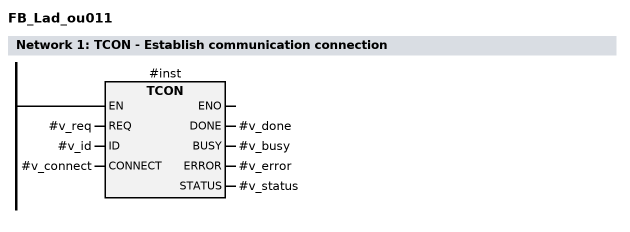
   #inst(REQ := #v_req,   // TCON
         ID := #v_id,
         CONNECT := #v_connect,
         DONE => #v_done,
         BUSY => #v_busy,
         ERROR => #v_error,
         STATUS => #v_status);
END_REGION
END_FUNCTION_BLOCK

FUNCTION_BLOCK "FB_Lad_ou012"   // FB78, LAD
{ S7_Optimized_Access := 'TRUE' }
   VAR_INPUT
      v_req : Bool;
      v_id : Word;
   END_VAR
   VAR_OUTPUT
      v_done : Bool;
      v_busy : Bool;
      v_error : Bool;
      v_status : Word;
   END_VAR
   VAR
      inst : TDISCON;
   END_VAR
BEGIN

REGION Network 1: TDISCON - Terminate communication connection
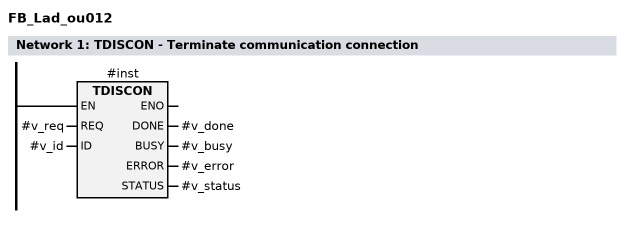
   #inst(REQ := #v_req, ID := #v_id, DONE => #v_done, BUSY => #v_busy, ERROR => #v_error, STATUS => #v_status);   // TDISCON
END_REGION
END_FUNCTION_BLOCK

FUNCTION_BLOCK "FB_Lad_ou013"   // FB79, LAD
{ S7_Optimized_Access := 'TRUE' }
   VAR_INPUT
      v_req : Bool;
      v_id : Conn_Ouc;
      v_len : UInt;
   END_VAR
   VAR_OUTPUT
      v_done : Bool;
      v_busy : Bool;
      v_error : Bool;
      v_status : Word;
   END_VAR
   VAR_IN_OUT
      v_data : Array[0..99] of Byte;
   END_VAR
   VAR
      inst : TSEND;
   END_VAR
BEGIN

REGION Network 1: TSEND - Send data via communication connection
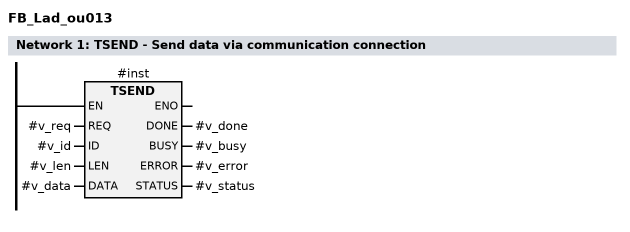
   #inst(REQ := #v_req,   // TSEND
         ID := #v_id,
         LEN := #v_len,
         DATA := #v_data,
         DONE => #v_done,
         BUSY => #v_busy,
         ERROR => #v_error,
         STATUS => #v_status);
END_REGION
END_FUNCTION_BLOCK

FUNCTION_BLOCK "FB_Lad_ou014"   // FB80, LAD
{ S7_Optimized_Access := 'TRUE' }
   VAR_INPUT
      v_req : Bool;
      v_id : Conn_Ouc;
      v_len : UDInt;
   END_VAR
   VAR_OUTPUT
      v_done : Bool;
      v_busy : Bool;
      v_error : Bool;
      v_status : Word;
   END_VAR
   VAR_IN_OUT
      v_data : Array[0..99] of Byte;
   END_VAR
   VAR
      inst : TSEND;
   END_VAR
BEGIN

REGION Network 1: TSEND - Send data via communication connection
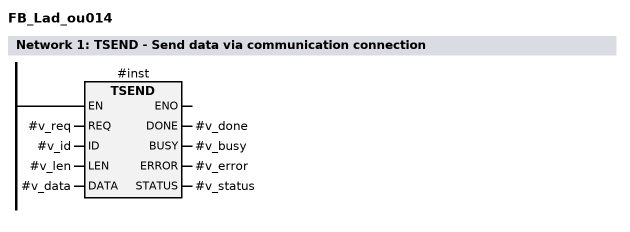
   #inst(REQ := #v_req,   // TSEND
         ID := #v_id,
         LEN := #v_len,
         DATA := #v_data,
         DONE => #v_done,
         BUSY => #v_busy,
         ERROR => #v_error,
         STATUS => #v_status);
END_REGION
END_FUNCTION_BLOCK

FUNCTION_BLOCK "FB_Lad_ou015"   // FB81, LAD
{ S7_Optimized_Access := 'TRUE' }
   VAR_INPUT
      v_en_r : Bool;
      v_id : Conn_Ouc;
      v_len : UInt;
      v_adhoc : Bool;
   END_VAR
   VAR_OUTPUT
      v_ndr : Bool;
      v_busy : Bool;
      v_error : Bool;
      v_status : Word;
      v_rcvd_len : UInt;
   END_VAR
   VAR_IN_OUT
      v_data : Array[0..99] of Byte;
   END_VAR
   VAR
      inst : TRCV;
   END_VAR
BEGIN

REGION Network 1: TRCV - Receive data via communication connection
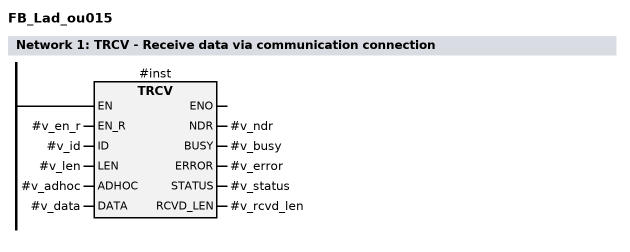
   #inst(EN_R := #v_en_r,   // TRCV
         ID := #v_id,
         LEN := #v_len,
         ADHOC := #v_adhoc,
         DATA := #v_data,
         NDR => #v_ndr,
         BUSY => #v_busy,
         ERROR => #v_error,
         STATUS => #v_status,
         RCVD_LEN => #v_rcvd_len);
END_REGION
END_FUNCTION_BLOCK

FUNCTION_BLOCK "FB_Lad_ou016"   // FB82, LAD
{ S7_Optimized_Access := 'TRUE' }
   VAR_INPUT
      v_en_r : Bool;
      v_id : Conn_Ouc;
      v_len : UDInt;
      v_adhoc : Bool;
   END_VAR
   VAR_OUTPUT
      v_ndr : Bool;
      v_busy : Bool;
      v_error : Bool;
      v_status : Word;
      v_rcvd_len : UDInt;
   END_VAR
   VAR_IN_OUT
      v_data : Array[0..99] of Byte;
   END_VAR
   VAR
      inst : TRCV;
   END_VAR
BEGIN

REGION Network 1: TRCV - Receive data via communication connection
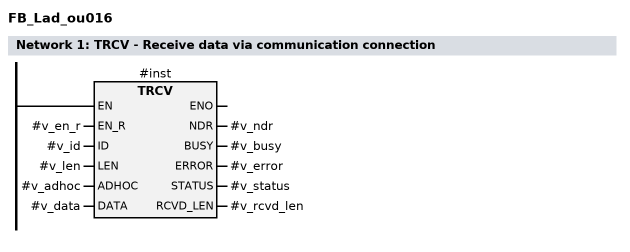
   #inst(EN_R := #v_en_r,   // TRCV
         ID := #v_id,
         LEN := #v_len,
         ADHOC := #v_adhoc,
         DATA := #v_data,
         NDR => #v_ndr,
         BUSY => #v_busy,
         ERROR => #v_error,
         STATUS => #v_status,
         RCVD_LEN => #v_rcvd_len);
END_REGION
END_FUNCTION_BLOCK

FUNCTION_BLOCK "FB_Lad_ou017"   // FB83, LAD
{ S7_Optimized_Access := 'TRUE' }
   VAR_INPUT
      v_req : Bool;
      v_id : Conn_Ouc;
      v_len : UDInt;
   END_VAR
   VAR_OUTPUT
      v_done : Bool;
      v_busy : Bool;
      v_error : Bool;
      v_status : Word;
   END_VAR
   VAR_IN_OUT
      v_data : Array[0..99] of Byte;
      v_addr : Array[0..99] of Byte;
   END_VAR
   VAR
      inst : TUSEND;
   END_VAR
BEGIN

REGION Network 1: TUSEND - Sending data
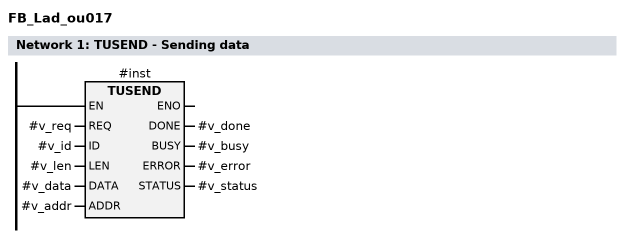
   #inst(REQ := #v_req,   // TUSEND
         ID := #v_id,
         LEN := #v_len,
         DATA := #v_data,
         ADDR := #v_addr,
         DONE => #v_done,
         BUSY => #v_busy,
         ERROR => #v_error,
         STATUS => #v_status);
END_REGION
END_FUNCTION_BLOCK

FUNCTION_BLOCK "FB_Lad_ou018"   // FB84, LAD
{ S7_Optimized_Access := 'TRUE' }
   VAR_INPUT
      v_en_r : Bool;
      v_id : Conn_Ouc;
      v_len : UDInt;
   END_VAR
   VAR_OUTPUT
      v_ndr : Bool;
      v_error : Bool;
      v_busy : Bool;
      v_status : Word;
      v_rcvd_len : UDInt;
   END_VAR
   VAR_IN_OUT
      v_data : Array[0..99] of Byte;
      v_addr : Array[0..99] of Byte;
   END_VAR
   VAR
      inst : TURCV;
   END_VAR
BEGIN

REGION Network 1: TURCV - Receiving data
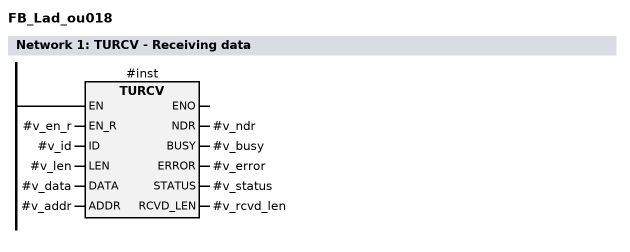
   #inst(EN_R := #v_en_r,   // TURCV
         ID := #v_id,
         LEN := #v_len,
         DATA := #v_data,
         ADDR := #v_addr,
         NDR => #v_ndr,
         BUSY => #v_busy,
         ERROR => #v_error,
         STATUS => #v_status,
         RCVD_LEN => #v_rcvd_len);
END_REGION
END_FUNCTION_BLOCK

FUNCTION_BLOCK "FB_Lad_ou019"   // FB85, LAD
{ S7_Optimized_Access := 'TRUE' }
   VAR_INPUT
      v_req : Bool;
      v_id : Conn_Ouc;
   END_VAR
   VAR_OUTPUT
      v_done : Bool;
      v_busy : Bool;
      v_error : Bool;
      v_status : Word;
   END_VAR
   VAR
      inst : T_RESET;
   END_VAR
BEGIN

REGION Network 1: T_RESET - Resetting the connection
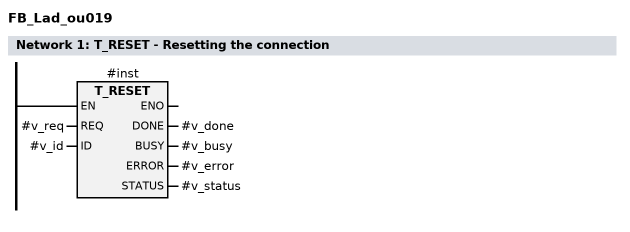
   #inst(REQ := #v_req, ID := #v_id, DONE => #v_done, BUSY => #v_busy, ERROR => #v_error, STATUS => #v_status);   // T_RESET
END_REGION
END_FUNCTION_BLOCK

FUNCTION_BLOCK "FB_Lad_ou020"   // FB86, LAD
{ S7_Optimized_Access := 'TRUE' }
   VAR_INPUT
      v_req : Bool;
      v_id : Word;
   END_VAR
   VAR_OUTPUT
      v_done : Bool;
      v_busy : Bool;
      v_error : Bool;
      v_status : Word;
   END_VAR
   VAR_IN_OUT
      v_result : Array[0..99] of Byte;
   END_VAR
   VAR
      inst : T_DIAG;
   END_VAR
BEGIN

REGION Network 1: T_DIAG - Checking the connection
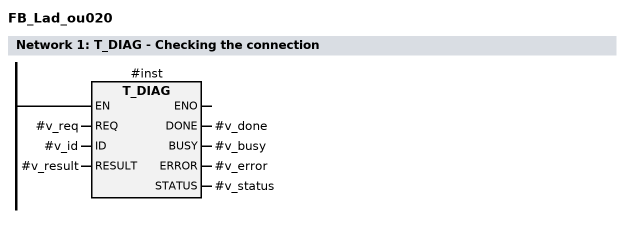
   #inst(REQ := #v_req,   // T_DIAG
         ID := #v_id,
         RESULT := #v_result,
         DONE => #v_done,
         BUSY => #v_busy,
         ERROR => #v_error,
         STATUS => #v_status);
END_REGION
END_FUNCTION_BLOCK

FUNCTION_BLOCK "FB_Lad_sc005"   // FB87, LAD
{ S7_Optimized_Access := 'TRUE' }
   VAR_INPUT
      v_req : Bool;
      v_r : Bool;
      v_id : Conn_Prg;
      v_r_id : Conn_R_Id;
   END_VAR
   VAR_OUTPUT
      v_done : Bool;
      v_error : Bool;
      v_status : Word;
   END_VAR
   VAR_IN_OUT
      v_sd_1 : Array[0..99] of Byte;
      v_len : Word;
   END_VAR
   VAR
      inst : BSEND;
   END_VAR
BEGIN

REGION Network 1: BSEND - Send data in segments
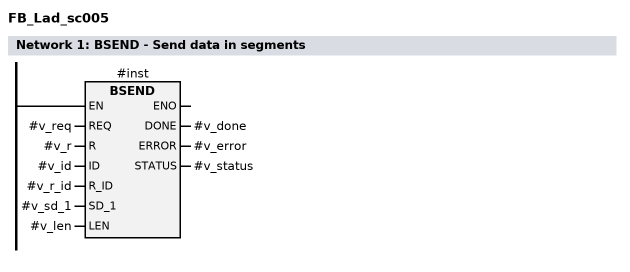
   #inst(REQ := #v_req,   // BSEND
         R := #v_r,
         ID := #v_id,
         R_ID := #v_r_id,
         SD_1 := #v_sd_1,
         LEN := #v_len,
         DONE => #v_done,
         ERROR => #v_error,
         STATUS => #v_status);
END_REGION
END_FUNCTION_BLOCK

FUNCTION_BLOCK "FB_Lad_sc006"   // FB88, LAD
{ S7_Optimized_Access := 'TRUE' }
   VAR_INPUT
      v_en_r : Bool;
      v_id : Conn_Prg;
      v_r_id : Conn_R_Id;
   END_VAR
   VAR_OUTPUT
      v_ndr : Bool;
      v_error : Bool;
      v_status : Word;
   END_VAR
   VAR_IN_OUT
      v_rd_1 : Array[0..99] of Byte;
      v_len : Word;
   END_VAR
   VAR
      inst : BRCV;
   END_VAR
BEGIN

REGION Network 1: BRCV - Receive data in segments
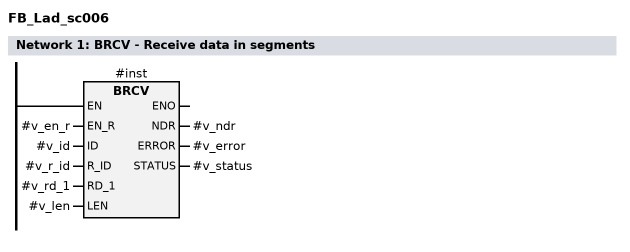
   #inst(EN_R := #v_en_r,   // BRCV
         ID := #v_id,
         R_ID := #v_r_id,
         RD_1 := #v_rd_1,
         LEN := #v_len,
         NDR => #v_ndr,
         ERROR => #v_error,
         STATUS => #v_status);
END_REGION
END_FUNCTION_BLOCK

FUNCTION_BLOCK "FB_Lad_ex011"   // FB89, LAD
{ S7_Optimized_Access := 'TRUE' }
VERSION : 0.1
   VAR_INPUT
      v_req : Bool;
      v_timezone : TimeTransformationRule;
   END_VAR
   VAR_OUTPUT
      v_done : Bool;
      v_busy : Bool;
      v_error : Bool;
      v_status : Word;
   END_VAR
   VAR
      inst : SET_TIMEZONE;
   END_VAR
BEGIN

REGION Network 1: SET_TIMEZONE - Set time zone
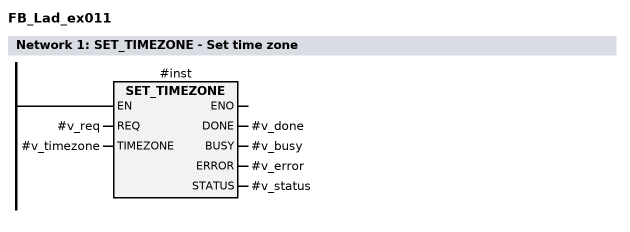
   #inst(REQ := #v_req,   // SET_TIMEZONE
         TimeZone := #v_timezone,
         DONE => #v_done,
         BUSY => #v_busy,
         ERROR => #v_error,
         STATUS => #v_status);
END_REGION
END_FUNCTION_BLOCK

FUNCTION_BLOCK "FB_Lad_ex045"   // FB90, LAD
{ S7_Optimized_Access := 'TRUE' }
   VAR_INPUT
      v_req : Bool;
      v_id : Hw_Io;
      v_index : DInt;
      v_mlen : UInt;
   END_VAR
   VAR_OUTPUT
      v_valid : Bool;
      v_busy : Bool;
      v_error : Bool;
      v_status : DWord;
      v_len : UInt;
   END_VAR
   VAR_IN_OUT
      v_record : Array[0..99] of Byte;
   END_VAR
   VAR
      inst : RDREC;
   END_VAR
BEGIN

REGION Network 1: RDREC - Read data record
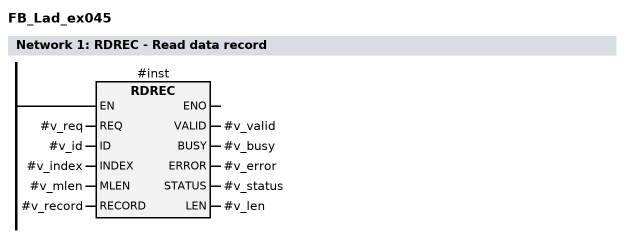
   #inst(REQ := #v_req,   // RDREC
         ID := #v_id,
         INDEX := #v_index,
         MLEN := #v_mlen,
         RECORD := #v_record,
         VALID => #v_valid,
         BUSY => #v_busy,
         ERROR => #v_error,
         STATUS => #v_status,
         LEN => #v_len);
END_REGION
END_FUNCTION_BLOCK

FUNCTION_BLOCK "FB_Lad_ex046"   // FB91, LAD
{ S7_Optimized_Access := 'TRUE' }
   VAR_INPUT
      v_req : Bool;
      v_id : Hw_Io;
      v_index : DInt;
      v_len : UInt;
   END_VAR
   VAR_OUTPUT
      v_done : Bool;
      v_busy : Bool;
      v_error : Bool;
      v_status : DWord;
   END_VAR
   VAR_IN_OUT
      v_record : Array[0..99] of Byte;
   END_VAR
   VAR
      inst : WRREC;
   END_VAR
BEGIN

REGION Network 1: WRREC - Write data record
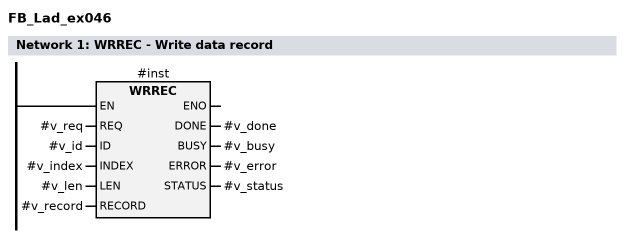
   #inst(REQ := #v_req,   // WRREC
         ID := #v_id,
         INDEX := #v_index,
         LEN := #v_len,
         RECORD := #v_record,
         DONE => #v_done,
         BUSY => #v_busy,
         ERROR => #v_error,
         STATUS => #v_status);
END_REGION
END_FUNCTION_BLOCK

FUNCTION_BLOCK "FB_Lad_ex047"   // FB92, LAD
{ S7_Optimized_Access := 'TRUE' }
   VAR_INPUT
      v_id : Hw_SubModule;
   END_VAR
   VAR_OUTPUT
      v_status : DWord;
      v_len : Int;
   END_VAR
   VAR_IN_OUT
      v_inputs : Array[0..99] of Byte;
   END_VAR
   VAR
      inst : GETIO;
   END_VAR
BEGIN

REGION Network 1: GETIO - Read all inputs of a submodule
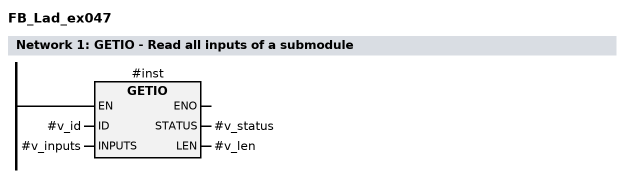
   #inst(ID := #v_id, INPUTS := #v_inputs, STATUS => #v_status, LEN => #v_len);   // GETIO
END_REGION
END_FUNCTION_BLOCK

FUNCTION_BLOCK "FB_Lad_ex048"   // FB93, LAD
{ S7_Optimized_Access := 'TRUE' }
   VAR_INPUT
      v_id : Hw_SubModule;
   END_VAR
   VAR_OUTPUT
      v_status : DWord;
   END_VAR
   VAR_IN_OUT
      v_outputs : Array[0..99] of Byte;
   END_VAR
   VAR
      inst : SETIO;
   END_VAR
BEGIN

REGION Network 1: SETIO - Write all outputs of a submodule
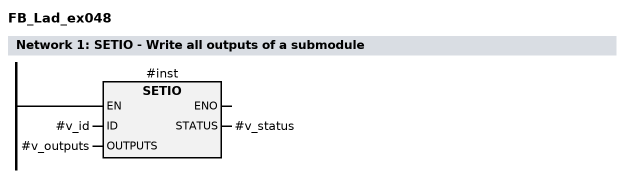
   #inst(ID := #v_id, OUTPUTS := #v_outputs, STATUS => #v_status);   // SETIO
END_REGION
END_FUNCTION_BLOCK

FUNCTION_BLOCK "FB_Lad_ex049"   // FB94, LAD
{ S7_Optimized_Access := 'TRUE' }
   VAR_INPUT
      v_id : Hw_SubModule;
      v_offset : Int;
      v_len : Int;
   END_VAR
   VAR_OUTPUT
      v_status : DWord;
      v_error : Bool;
   END_VAR
   VAR_IN_OUT
      v_inputs : Array[0..99] of Byte;
   END_VAR
   VAR
      inst : GETIO_PART;
   END_VAR
BEGIN

REGION Network 1: GETIO_PART - Read inputs of a submodule
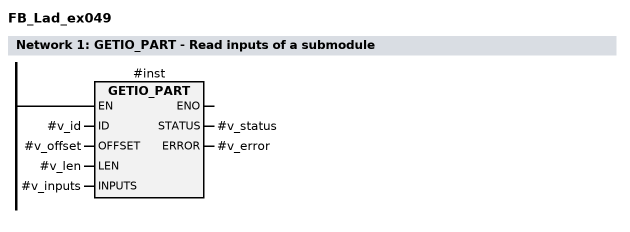
   #inst(ID := #v_id,   // GETIO_PART
         OFFSET := #v_offset,
         LEN := #v_len,
         INPUTS := #v_inputs,
         STATUS => #v_status,
         ERROR => #v_error);
END_REGION
END_FUNCTION_BLOCK

FUNCTION_BLOCK "FB_Lad_ex050"   // FB95, LAD
{ S7_Optimized_Access := 'TRUE' }
   VAR_INPUT
      v_id : Hw_SubModule;
      v_offset : Int;
      v_len : Int;
   END_VAR
   VAR_OUTPUT
      v_status : DWord;
      v_error : Bool;
   END_VAR
   VAR_IN_OUT
      v_outputs : Array[0..99] of Byte;
   END_VAR
   VAR
      inst : SETIO_PART;
   END_VAR
BEGIN

REGION Network 1: SETIO_PART - Write outputs of a submodule
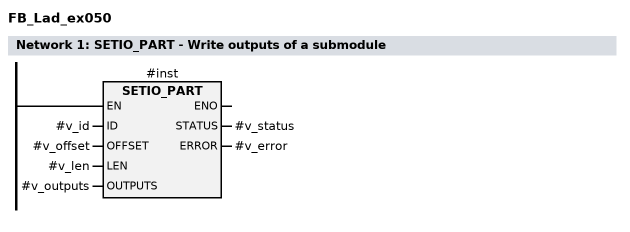
   #inst(ID := #v_id,   // SETIO_PART
         OFFSET := #v_offset,
         LEN := #v_len,
         OUTPUTS := #v_outputs,
         STATUS => #v_status,
         ERROR => #v_error);
END_REGION
END_FUNCTION_BLOCK

FUNCTION_BLOCK "FB_Lad_ex057"   // FB96, LAD
{ S7_Optimized_Access := 'TRUE' }
   VAR_INPUT
      v_req : Bool;
      v_mode : UInt;
      v_laddr : Hw_Interface;
      v_ctrlrec : Array[0..99] of Byte;
   END_VAR
   VAR_OUTPUT
      v_done : Bool;
      v_busy : Bool;
      v_error : Bool;
      v_status : DWord;
      v_err_info : Word;
   END_VAR
   VAR
      inst : ReconfigIOSystem;
   END_VAR
BEGIN

REGION Network 1: ReconfigIOSystem - Reconfigure IO system
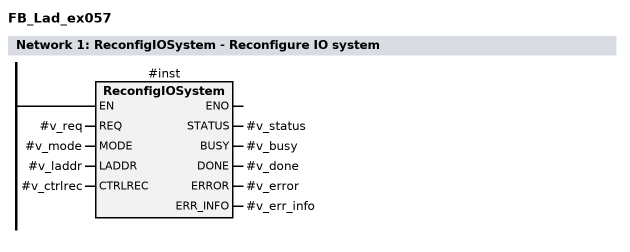
   #inst(REQ := #v_req,   // ReconfigIOSystem
         MODE := #v_mode,
         LADDR := #v_laddr,
         CTRLREC := #v_ctrlrec,
         STATUS => #v_status,
         BUSY => #v_busy,
         DONE => #v_done,
         ERROR => #v_error,
         ERR_INFO => #v_err_info);
END_REGION
END_FUNCTION_BLOCK

FUNCTION_BLOCK "FB_Lad_ex062"   // FB97, LAD
{ S7_Optimized_Access := 'TRUE' }
   VAR_INPUT
      v_mode : Int;
      v_f_id : Hw_SubModule;
      v_mlen : Int;
      v_code1 : Byte;
      v_code2 : Byte;
   END_VAR
   VAR_OUTPUT
      v_new : Bool;
      v_status : DWord;
      v_slot : Hw_SubModule;
      v_subslot : Hw_SubModule;
      v_index : UInt;
      v_len : UInt;
   END_VAR
   VAR_IN_OUT
      v_record : Array[0..99] of Byte;
   END_VAR
   VAR
      inst : RCVREC;
   END_VAR
BEGIN

REGION Network 1: RCVREC - Receive data record
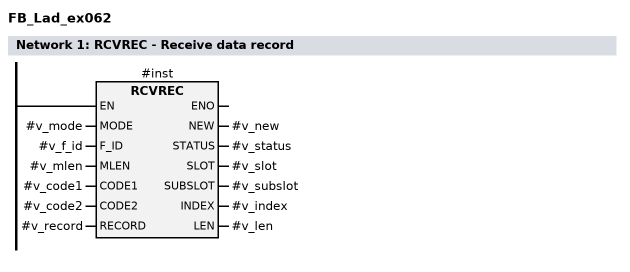
   #inst(MODE := #v_mode,   // RCVREC
         F_ID := #v_f_id,
         MLEN := #v_mlen,
         CODE1 := #v_code1,
         CODE2 := #v_code2,
         RECORD := #v_record,
         NEW => #v_new,
         STATUS => #v_status,
         SLOT => #v_slot,
         SUBSLOT => #v_subslot,
         INDEX => #v_index,
         LEN => #v_len);
END_REGION
END_FUNCTION_BLOCK

FUNCTION_BLOCK "FB_Lad_ex063"   // FB98, LAD
{ S7_Optimized_Access := 'TRUE' }
   VAR_INPUT
      v_mode : Int;
      v_f_id : Hw_SubModule;
      v_code1 : Byte;
      v_code2 : Byte;
      v_len : UInt;
   END_VAR
   VAR_OUTPUT
      v_new : Bool;
      v_status : DWord;
      v_slot : Hw_SubModule;
      v_subslot : Hw_SubModule;
      v_index : UInt;
      v_rlen : UInt;
   END_VAR
   VAR_IN_OUT
      v_record : Array[0..99] of Byte;
   END_VAR
   VAR
      inst : PRVREC;
   END_VAR
BEGIN

REGION Network 1: PRVREC - Make data record available
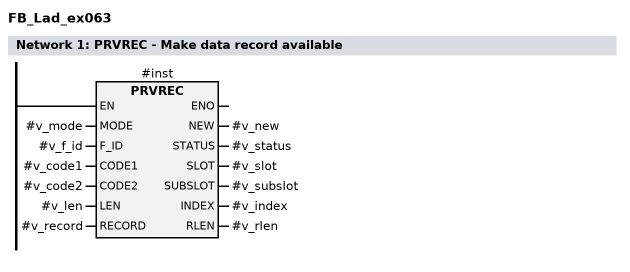
   #inst(MODE := #v_mode,   // PRVREC
         F_ID := #v_f_id,
         CODE1 := #v_code1,
         CODE2 := #v_code2,
         LEN := #v_len,
         RECORD := #v_record,
         NEW => #v_new,
         STATUS => #v_status,
         SLOT => #v_slot,
         SUBSLOT => #v_subslot,
         INDEX => #v_index,
         RLEN => #v_rlen);
END_REGION
END_FUNCTION_BLOCK

FUNCTION_BLOCK "FB_Lad_ex096"   // FB99, LAD
{ S7_Optimized_Access := 'TRUE' }
   VAR_INPUT
      v_req : Bool;
      v_laddr : Hw_Io;
      v_index : Int;
   END_VAR
   VAR_OUTPUT
      v_valid : Bool;
      v_busy : Bool;
      v_error : Bool;
      v_status : DWord;
      v_len : Int;
   END_VAR
   VAR_IN_OUT
      v_record : Array[0..99] of Byte;
   END_VAR
   VAR
      inst : RD_DPAR;
   END_VAR
BEGIN

REGION Network 1: RD_DPAR - Read module data record
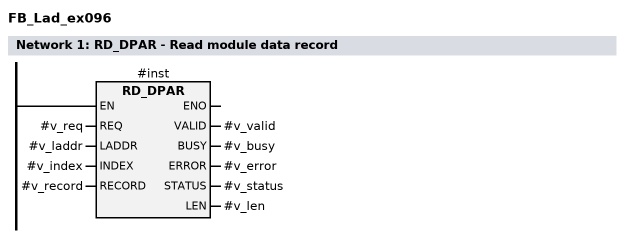
   #inst(REQ := #v_req,   // RD_DPAR
         LADDR := #v_laddr,
         INDEX := #v_index,
         RECORD := #v_record,
         VALID => #v_valid,
         BUSY => #v_busy,
         ERROR => #v_error,
         STATUS => #v_status,
         LEN => #v_len);
END_REGION
END_FUNCTION_BLOCK

FUNCTION_BLOCK "FB_Lad_ex127"   // FB100, LAD
{ S7_Optimized_Access := 'TRUE' }
   VAR_INPUT
      v_laddr : Hw_Io;
      v_im_type : UInt;
   END_VAR
   VAR_OUTPUT
      v_done : Bool;
      v_busy : Bool;
      v_error : Bool;
      v_status : Word;
   END_VAR
   VAR_IN_OUT
      v_data : Array[0..99] of Byte;
   END_VAR
   VAR
      inst : Get_IM_Data;
   END_VAR
BEGIN

REGION Network 1: Get_IM_Data - Reading identification and maintenance data
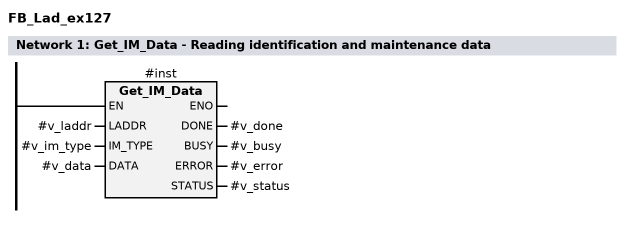
   #inst(LADDR := #v_laddr,   // Get_IM_Data
         IM_TYPE := #v_im_type,
         DATA := #v_data,
         DONE => #v_done,
         BUSY => #v_busy,
         ERROR => #v_error,
         STATUS => #v_status);
END_REGION
END_FUNCTION_BLOCK

FUNCTION_BLOCK "FB_Lad_ex128"   // FB101, LAD
{ S7_Optimized_Access := 'TRUE' }
   VAR_INPUT
      v_laddr : Hw_IoSystem;
      v_station_nr : UInt;
   END_VAR
   VAR_OUTPUT
      v_done : Bool;
      v_busy : Bool;
      v_error : Bool;
      v_len : DInt;
      v_status : Word;
   END_VAR
   VAR_IN_OUT
      v_data : Array[0..99] of Byte;
   END_VAR
   VAR
      inst : Get_Name;
   END_VAR
BEGIN

REGION Network 1: GET_NAME - Read out name of an IO device or a DP slave
